(*
SPDX-FileCopyrightText: c 2026 Oleksandr Tiutyk <trofimich@gmail.com>
SPDX-License-Identifier: MIT
License: https://opensource.org/license/mit
*)

(*!
<summary>Groups the four cyclic file-content manager scenarios.</summary>
<description>
Owns one independent directory fixture per leaf. Each child borrows and exclusively drives its assigned fixture.
The group keeps the fixtures, Children array and parent associations fixed for the lifetime of the tests.
Use from one task without reentry. Do not copy the group or modify its borrowed Children array.
</description>
*)

{attribute 'no_assign'}
{attribute 'no_explicit_call' := 'do not call this function block directly'}
FUNCTION_BLOCK FileContentManagerOperationsTest EXTENDS TOF_Testing.TestGroup<4>
VAR_STAT
	//! <summary>Class name shared by instances of this concrete function block.</summary>
	{attribute 'hide'}
	_ClassName : STRING := __POUNAME();
END_VAR
VAR
	_TextDirectory : FileTestDirectory(directoryPath := 'C:\OpenFrameworkTests\FileContent_CreateText');
	_ReadOnlyDirectory : FileTestDirectory(directoryPath := 'C:\OpenFrameworkTests\FileContent_ReadOnly');
	_CancelDirectory : FileTestDirectory(directoryPath := 'C:\OpenFrameworkTests\FileContent_Cancel');
	_ReuseDirectory : FileTestDirectory(directoryPath := 'C:\OpenFrameworkTests\FileContent_Reuse');

	_TextTest : FileTextReadWriteTest(
		name := "CreateTextFile",
		parent := THIS^,
		directory := _TextDirectory,
		scenarioTimeout := T#10S
	);
	_ReadOnlyTest : FileReadOnlyWriteTest(
		name := "WriteToFileOpenedForReading",
		parent := THIS^,
		directory := _ReadOnlyDirectory,
		scenarioTimeout := T#15S
	);
	_CancelTest : FileWriteCancellationTest(
		name := "CancelDuringFileWrite",
		parent := THIS^,
		directory := _CancelDirectory,
		scenarioTimeout := T#10S
	);
	_ReuseTest : FileManagerReuseTest(
		name := "ReuseAfterReset",
		parent := THIS^,
		directory := _ReuseDirectory,
		scenarioTimeout := T#20S
	);

	_Children : ARRAY [0.._ChildCount - 1] OF TOF_Testing.ITestElement :=
	[
		_TextTest,
		_ReadOnlyTest,
		_CancelTest,
		_ReuseTest
	];
END_VAR

//! <summary>Borrows the fixed leaf array for this group's lifetime; callers must not modify it.</summary>
{attribute 'monitoring' := 'call'}
PROPERTY Children : REFERENCE TO ARRAY [0.._ChildCount - 1] OF TOF_Testing.ITestElement
GET
Children REF= _Children;
END_GET
END_PROPERTY

//! <summary>Borrows this concrete type name; callers must not modify the referenced storage.</summary>
{attribute 'monitoring' := 'call'}
PROPERTY ClassName : REFERENCE TO STRING
GET
ClassName REF= _ClassName;
END_GET
END_PROPERTY

//! <summary>Borrows the compiler-initialized namespace; callers must not modify the returned reference.</summary>
{attribute 'monitoring' := 'call'}
PROPERTY NamespaceName : REFERENCE TO STRING
GET
NamespaceName REF= CurrentNamespace.Name;
END_GET
END_PROPERTY

//! <summary>Reports this concrete instance size, excluding separately allocated storage.</summary>
{attribute 'monitoring' := 'call'}
PROPERTY SelfSize : ULINT
GET
SelfSize := XSIZEOF(THIS^);
END_GET
END_PROPERTY

END_FUNCTION_BLOCK

(* stored: Version 1.1.0.1
   POU FileContentManagerOperationsTest: Id {38864847-5983-433d-a770-6ea5c772c1a2}, SpecialFunc None
   Property Children: Id {53679131-82c1-4520-958b-a4126e5547c4}
   Get Get: Id {bdbebcf2-368c-4b32-86ce-1b80b2096fe6}
   Property ClassName: Id {0e328233-4437-4ba7-9929-6ddc7a423ba1}
   Get Get: Id {05c6e581-0b64-4875-ae64-7f0ffa202a1c}
   Property NamespaceName: Id {f8c4819c-e034-43af-aa3a-0de302692ebd}
   Get Get: Id {3e4f788d-f206-4f9b-a08b-d381f553f2c8}
   Property SelfSize: Id {d9ee4ad6-4b0f-4f4b-9349-9bb9eecb1987}
   Get Get: Id {d0caaa54-f989-4627-96df-3505e5714b74} *)
